// TIA Portal V21 export
// export: Created 2026-10-23T21:22:26.9798531Z, ExportSetting WithReadOnly, DisplayName Totally Integrated Automation Portal, DisplayVersion V21 Update 1, DisplayName SINAMICS Startdrive Advanced, DisplayVersion V21 HF2, DisplayName SINAMICS Startdrive G110M, G120, G120C, G120D, G120P, G115D, DisplayVersion V21 HF2, DisplayName SINAMICS Startdrive G130, G150, S120, S150, G200, G220, S200, S210, S220, Innomotics MVD, DisplayVersion V21 HF2, DisplayName STEP 7 Professional, DisplayVersion V21 Update 1, DisplayName STEP 7 Safety, DisplayVersion V21, DisplayName Tech WebApplication, DisplayVersion V21, DisplayName WinCC Basic/Comfort/Advanced, DisplayVersion V21 Update 1, DisplayName WinCC Unified, DisplayVersion V21 Update 1
ORGANIZATION_BLOCK "OB_Main"   // OB1, SCL, ProgramCycle
TITLE = "Main Program Sweep (Cycle)" / Main program of PLC_1200
{ S7_Optimized_Access := 'TRUE' }
// Calls the conveyor with the onboard inputs and output of the CPU 1214C
// stored: CodeModifiedDate 2026-10-23T19:59:16.3446293Z, CompileDate 2026-10-23T19:59:16.3446293Z, ConstantName OB_OB_Main, CreationDate 2026-10-23T19:59:09.2129607Z, DownloadDate 0001-01-01T00:00:00Z, EventClass Program cycle, InterfaceModifiedDate 2008-07-21T16:55:08.419547Z, IsConsistent true, LoadMemoryLength 4275, ModifiedDate 2026-10-23T19:59:16.3446293Z, ParameterModified 2008-07-21T16:55:08.419547Z, PriorityNumber 1, ProcessImagePartNumber 65535, SetENOAutomatically false, StructureModified 2008-07-21T16:55:08.419547Z, WorkMemoryLength 88
   VAR_INPUT
      Initial_Call : Bool;   // Initial call of this OB
      Remanence : Bool;   // =True, if remanent data are available
   END_VAR
BEGIN

       REGION Conveyor
           "IDB_Conveyor1200"(Start := "BeltStart",
                              Stop := "BeltStop",
                              SpeedRaw := "BeltSpeedRaw",
                              Motor => "BeltMotor");
       END_REGION
END_ORGANIZATION_BLOCK
